FUNCTION_BLOCK FB_SFC_Template EXTENDS FB_SFC_Cycle IMPLEMENTS ITF_FB_SFC_Cycle
VAR_INPUT
END_VAR
VAR_OUTPUT
END_VAR
VAR
END_VAR

m_Set_SFCFlags_Reference();
SUPER^();

ACTION act_Oper:
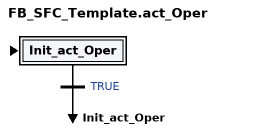
INITIAL_STEP Init_act_Oper:
END_STEP
TRANSITION FROM Init_act_Oper TO Init_act_Oper
    := TRUE;
END_TRANSITION
END_ACTION

METHOD m_Set_SFCFlags_Reference : BOOL
//Set reference to SFC flags

refSFC.SFCInit REF= SFCInit;
refSFC.SFCReset REF= SFCReset;
refSFC.SFCError REF= SFCError;
refSFC.SFCEnableLimit REF= SFCEnableLimit;
refSFC.SFCErrorStep REF= SFCErrorStep;
refSFC.SFCErrorPOU REF= SFCErrorPOU;
refSFC.SFCQuitError REF= SFCQuitError;
refSFC.SFCPause REF= SFCPause;
refSFC.SFCTrans REF= SFCTrans;
refSFC.SFCCurrentStep REF= SFCCurrentStep;
refSFC.SFCTip REF= SFCTip;
refSFC.SFCTipMode REF= SFCTipMode;

// Cycle handle for SFC
m_SFC_Handle();
END_METHOD

END_FUNCTION_BLOCK

(* stored: Version 1.1.0.1, ProductVersion 3.1.4024.12
   POU FB_SFC_Template: Id {03ecb4ba-29f7-4048-a93a-8d5c53cd05cb}, SpecialFunc None
   Action act_Oper: Id {04ae6814-7809-4820-9c1c-a19561775a17}
   Method m_Set_SFCFlags_Reference: Id {4cf88e6d-ae8b-4924-927c-6335e6620f0b} *)
